// TIA Portal V17 export
DATA_BLOCK "MCP_RC_DB4"   // DB9804
{ S7_Optimized_Access := 'TRUE' }
   VAR
      "A" : "MCP_RC_UDT";
      "B" : "MCP_RC_UDT";
   END_VAR
BEGIN
END_DATA_BLOCK
